Staubli VAL3: getPointIndex.pgx

public program getPointIndex(string x_sTrajItem, string x_sPoint, num& x_nPointIndex, bool& x_bResult)
  local bool l_bResult
  local num l_nSize
begin
  toNum(x_sPoint,x_nPointIndex,x_bResult)
  if !x_bResult
    call getPointSize(x_sTrajItem,l_nSize)
    x_nPointIndex=l_nSize-1
  endIf
end
